(* IEC 61131-3 sources: llm-plc-st-eval/data/processed_definitivo/gemini-3.1-pro-preview/I6/few_shot, 3 files *)

(* ---- ejec_1.st ---- *)
FUNCTION_BLOCK FB_Temperatura
VAR_INPUT
    rawTemp : INT; (* Valor crudo del sensor (0-27648) *)
END_VAR
VAR_OUTPUT
    tempC : REAL; (* Temperatura en grados Celsius (0.0-100.0) *)
    enfriador : BOOL; (* Estado del enfriador *)
    almSensor : BOOL; (* Alarma de sensor fuera de rango *)
END_VAR

(* Evaluacion de limites para la alarma del sensor *)
almSensor := (rawTemp < 0) OR (rawTemp > 27648);

(* Escalado de la señal analogica *)
tempC := INT_TO_REAL(rawTemp) * 100.0 / 27648.0;

(* Control del enfriador con histeresis y proteccion por alarma *)
IF almSensor THEN
    enfriador := FALSE;
ELSIF tempC >= 80.0 THEN
    enfriador := TRUE;
ELSIF tempC <= 75.0 THEN
    enfriador := FALSE;
END_IF;
END_FUNCTION_BLOCK

(* ---- ejec_2.st ---- *)
FUNCTION_BLOCK FB_Temperatura
VAR_INPUT
    rawTemp : INT; (* Valor crudo del sensor de temperatura *)
END_VAR
VAR_OUTPUT
    tempC : REAL; (* Temperatura escalada en grados Celsius *)
    enfriador : BOOL; (* Estado del enfriador *)
    almSensor : BOOL; (* Alarma de sensor fuera de rango *)
END_VAR

(* Calculo de la temperatura escalada (0.0 a 100.0) *)
tempC := (INT_TO_REAL(rawTemp) / 27648.0) * 100.0;

(* Evaluacion de alarma por limites del sensor *)
almSensor := (rawTemp < 0) OR (rawTemp > 27648);

(* Control del enfriador con histeresis y bloqueo por alarma *)
IF almSensor THEN
    enfriador := FALSE;
ELSIF tempC >= 80.0 THEN
    enfriador := TRUE;
ELSIF tempC <= 75.0 THEN
    enfriador := FALSE;
END_IF;
END_FUNCTION_BLOCK

(* ---- ejec_3.st ---- *)
FUNCTION_BLOCK FB_Temperatura
VAR_INPUT
    rawTemp : INT; (* Valor crudo del sensor de temperatura *)
END_VAR
VAR_OUTPUT
    tempC : REAL; (* Temperatura calculada en grados Celsius *)
    enfriador : BOOL; (* Señal de activacion del enfriador *)
    almSensor : BOOL; (* Alarma de sensor fuera de rango *)
END_VAR

(* Deteccion de falla o fuera de rango del sensor *)
almSensor := (rawTemp < 0) OR (rawTemp > 27648);

(* Acondicionamiento y escalado de la señal (0-27648 a 0.0-100.0) *)
tempC := (INT_TO_REAL(rawTemp) / 27648.0) * 100.0;

(* Control del enfriador con histeresis y proteccion por alarma *)
IF almSensor THEN
    enfriador := FALSE; (* Apaga el enfriador si hay error en el sensor *)
ELSE
    IF tempC >= 80.0 THEN
        enfriador := TRUE; (* Activa por alta temperatura *)
    ELSIF tempC <= 75.0 THEN
        enfriador := FALSE; (* Desactiva al alcanzar el umbral inferior *)
    END_IF;
    (* Entre 75.0 y 80.0 conserva su estado anterior *)
END_IF;
END_FUNCTION_BLOCK
